FUNCTION FC 1 : VOID
BEGIN
NETWORK
      A I 0.0 I 0.1
END_FUNCTION
